DATA_BLOCK "FRK_LineSetStage"
{ S7_Optimized_Access := 'TRUE' }
VERSION : 0.1
NON_RETAIN
VAR
    Values {ExternalAccessible := 'False'; ExternalVisible := 'False'; ExternalWritable := 'False'} : "ST_LineProbeConfig";
END_VAR
BEGIN
END_DATA_BLOCK
